// TIA Portal V20 export
// export: Created 2026-10-12T16:46:22.6670983Z, ExportSetting WithDefaults, DisplayName Totally Integrated Automation Portal, DisplayVersion V20 Update 6, DisplayName TIA Portal Openness, DisplayVersion V20 Update 6, DisplayName TIA Portal Version Control Interface, DisplayVersion V20 Update 6, DisplayName SINAMICS Startdrive Advanced, DisplayVersion V20 SP1 Update 2, DisplayName SINAMICS Startdrive G110M, G120, G120C, G120D, G120P, G115D, DisplayVersion V20 SP1 Update 2, DisplayName SINAMICS Startdrive G130, G150, S120, S150, SINAMICS MV, G220, S200, S210, DisplayVersion V20 SP1 Update 2, DisplayName STEP 7 Professional, DisplayVersion V20 Update 6, DisplayName STEP 7 Safety, DisplayVersion V20 Update 2, DisplayName WinCC Basic/Comfort/Advanced, DisplayVersion V20 Update 6, DisplayName WinCC Professional, DisplayVersion V20 Update 6, DisplayName WinCC Unified, DisplayVersion V20 Update 6
TYPE "UDT_Artikel"
// stored: IsFailsafeCompliant false
   STRUCT
      ID : Int;
      "Name" : String;
      Beschreibung : String;
      Aktiv : Bool;
      SAP_Nummer : String;
      Kunde : String;
      Prozess : String;
      Zeichnungsnummer : Int;
      Prozessfreigabe_Datum : Date_And_Time;
      Prozessfreigabe_Name : String;
      Freitext_1 : String;
      Freitext_2 : String;
      Freitext_3 : String;
   END_STRUCT;
END_TYPE
